Staubli VAL3: setDigOutput.pgx

public program setDigOutput(num x_nIndex, bool x_bValue, num& x_nResult)
  local string l_sDesc
  local string l_sPath
//写数字输出 dOutput[x_nIndex]
//返回码 x_nResult: 0=正常  -1=索引越界  -2=该位未绑定物理通道(ioStatus<0，写入无效)
//注意：dOutput 还没有 link（未做物理 IO 导入），此时写入不会作用到任何物理点，
//      必须先在 SRS 里完成物理 IO 导入，见 docs/05-IO绑定方法.md
begin
  x_nResult=0

  //越界检查：合法下标 0..size(dOutput)-1（手册 2.5.4，第31页 num size(*)）
  if (x_nIndex<0) or (x_nIndex>=size(dOutput))
    x_nResult=-1
    return
  endIf

  //未绑定物理通道时先拦截：手册 3.5.2（第59页）——给未 link 的 dio 赋值会触发 runtime error
  if ioStatus(dOutput[x_nIndex],l_sDesc,l_sPath)<0
    x_nResult=-2
    return
  endIf

  dOutput[x_nIndex]=x_bValue
end
